(* IEC 61131-3 sources: plcassist-cli/packages/volt-lsp-iec/test-corpus/pro2193/Device/Plc Logic/Application/03 Hardware Units/31 SER/31.02 - X Units/Xi Unit in project, 2 files *)

(* ---- IXiUnit_Commands.itf ---- *)
// Commands specific for an Xu Unit
INTERFACE IXiUnit_Commands

END_INTERFACE

(* ---- XiUnitFB.fb ---- *)
{attribute 'symbol' := 'none'}
FUNCTION_BLOCK XiUnitFB
EXTENDS XiUnit_DefaultFB
IMPLEMENTS IXiUnit_Commands
VAR_INPUT
END_VAR
VAR_IN_OUT
	DataProject					: XiUnit_Data;
END_VAR
VAR
END_VAR

SUPER^(
	Data				:= Data,
	AxisRef				:= AxisRef,
	DataBrink			:= DataBrink,
	coveredDistance		:= coveredDistance,
);

END_FUNCTION_BLOCK
